// TIA Portal V20 export
TYPE "T2_UDT_Padre"
// Prueba IA 2: UDT con UDT anidado y array
   STRUCT
      Id : DInt;   // Identificador
      Hijo : "T2_UDT_Hijo";   // UDT anidado
      Lista : Array[0..3] of Int;   // Array dentro de UDT
      Activo : Bool;   // Bit
   END_STRUCT;
END_TYPE
